SUBAPPLICATION Uebung_141_AX (* Übung zu DiagSetDTC: Drahtbruch 4-20 mA als DTC über DM1 *)
  (* Standard: 61499-2; Description: Copyright (c) 2026 Meisterschulen am Ostbahnhof This program and the accompanying materials are made available under the terms of the Eclipse Public License 2.0 which is available at https://www.eclipse.org/legal/epl-2.0/ SPDX-License-Identifier: EPL-2.0 *)
  (* Version 1.0, 2026-11-17, Franz Höpfinger, Meisterschulen am Ostbahnhof, initial API and implementation and/or initial documentation *)
  PACKAGE Uebungen;
  IMPORT Uebungen::const::Uebung_120_129::Filter::ADD_ALL_PASS;
  IMPORT Uebungen::const::Uebung_120_129::Filter::FLT_ALL_PASS;
  IMPORT Uebungen::const::Uebung_140_149::Diag::MV_DRAHTBRUCH;
  IMPORT Uebungen::const::Uebung_140_149::Diag::MV_OK;
  IMPORT Uebungen::const::Uebung_140_149::Diag::SPN_DRAHTBRUCH_AI6;
  IMPORT isobus::pgn::ISOUSERHOME_e::thisMember;
  IMPORT isobus::pgn::ISO_CAN_NODE::NODE1;
  IMPORT isobus::pgn::diag::FMI::CURRENT_LOW_OPEN_CIRCUIT;
  IMPORT logiBUS::io::AI::logiBUS_AI::AnalogInput_I6;
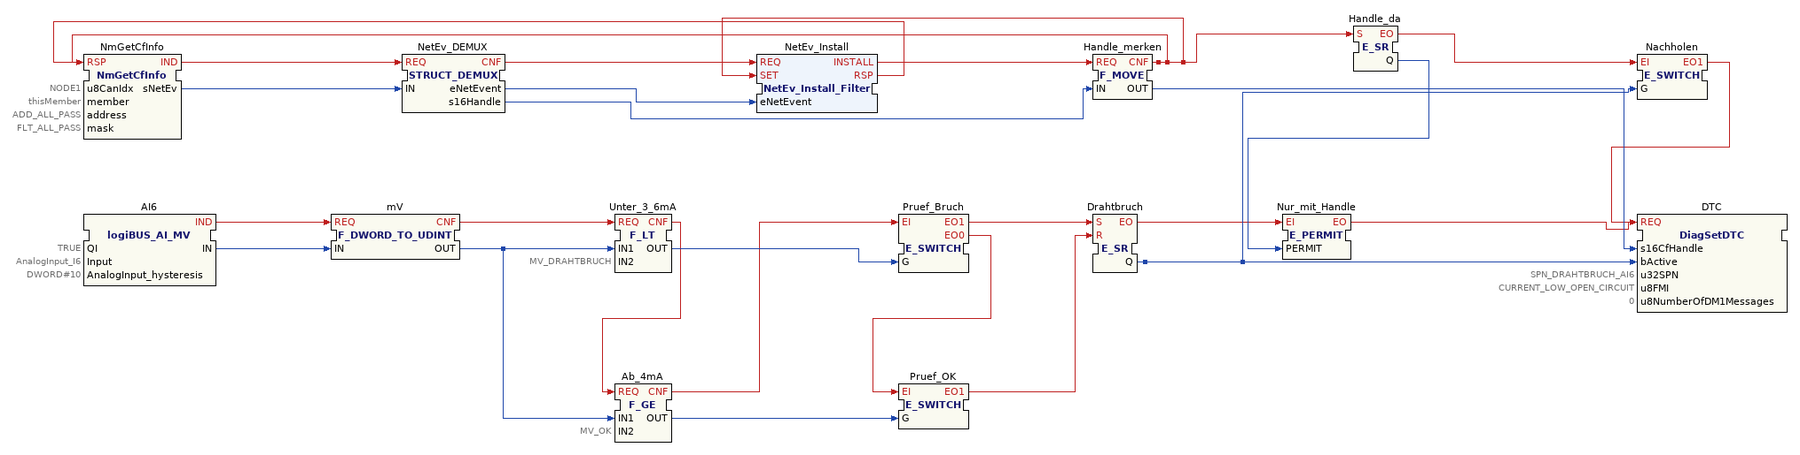
  (* Drahtbruch 4-20 mA an AI6 als DTC über DM1 (DiagSetDTC) Pin-mV unter 564 (3,6 mA) = Drahtbruch, wieder OK ab 626 (4 mA). Eigener CF-Handle aus NmGetCfInfo (thisMember, Active/NewAddress), RSP immer. DTC nur bei Zustandswechsel: SPN 520192, FMI 5, aktiv bis gelöscht. Test: Kabel ab = DM1 mit SPN 520192/FMI 5, jede Sekunde. Kabel dran = DTC inaktiv, in DM2, mit DM3 löschbar. Braucht Firmware ab LOGIBUS 96f591f2 (DM1) und isobus_pgn-ELF mit DiagSetDTC. *)
  FBS
    NmGetCfInfo : isobus::pgn::NmGetCfInfo(u8CanIdx := NODE1, member := thisMember, address := ADD_ALL_PASS, mask := FLT_ALL_PASS);
    NetEv_DEMUX : eclipse4diac::convert::STRUCT_DEMUX; {SET_ATTRIBUTE(StructuredType, isobus::pgn::ISONETEVENT_T)}
    Handle_merken : iec61131::selection::F_MOVE; (* eigener CF-Handle (s16Handle) *)
    Handle_da : iec61499::events::E_SR;
    Nachholen : iec61499::events::E_SWITCH; (* Drahtbruch schon vor dem Handle da: jetzt melden *)
    AI6 : logiBUS::io::AI::logiBUS_AI_MV(QI := TRUE, Input := AnalogInput_I6, AnalogInput_hysteresis := DWORD#10); (* mV am Pin, 4-20 mA über 491,2 Ohm *)
    mV : iec61131::conversion::F_DWORD_TO_UDINT;
    Unter_3_6mA : iec61131::comparison::F_LT(IN2 := MV_DRAHTBRUCH);
    Ab_4mA : iec61131::comparison::F_GE(IN2 := MV_OK);
    Pruef_Bruch : iec61499::events::E_SWITCH;
    Pruef_OK : iec61499::events::E_SWITCH;
    Drahtbruch : iec61499::events::E_SR; (* EO nur bei Zustandswechsel *)
    Nur_mit_Handle : iec61499::events::E_PERMIT;
    DTC : isobus::pgn::diag::DiagSetDTC(u32SPN := SPN_DRAHTBRUCH_AI6, u8FMI := CURRENT_LOW_OPEN_CIRCUIT, u8NumberOfDM1Messages := 0); (* DM1: SPN 520192, FMI 5 *)
  END_FBS
  SUBAPPS
    NetEv_Install : MyLib::sys::NetEv_Install_Filter;
  END_SUBAPPS
  EVENT_CONNECTIONS
    NmGetCfInfo.IND TO NetEv_DEMUX.REQ;
    NetEv_DEMUX.CNF TO NetEv_Install.REQ;
    NetEv_Install.INSTALL TO Handle_merken.REQ;
    NetEv_Install.RSP TO NmGetCfInfo.RSP;
    Handle_merken.CNF TO NetEv_Install.SET;
    Handle_merken.CNF TO Handle_da.S;
    Handle_merken.CNF TO NmGetCfInfo.RSP;
    Handle_da.EO TO Nachholen.EI;
    Nachholen.EO1 TO DTC.REQ;
    AI6.IND TO mV.REQ;
    mV.CNF TO Unter_3_6mA.REQ;
    Unter_3_6mA.CNF TO Ab_4mA.REQ;
    Ab_4mA.CNF TO Pruef_Bruch.EI;
    Pruef_Bruch.EO1 TO Drahtbruch.S;
    Pruef_Bruch.EO0 TO Pruef_OK.EI;
    Pruef_OK.EO1 TO Drahtbruch.R;
    Drahtbruch.EO TO Nur_mit_Handle.EI;
    Nur_mit_Handle.EO TO DTC.REQ;
  END_CONNECTIONS
  DATA_CONNECTIONS
    NmGetCfInfo.sNetEv TO NetEv_DEMUX.IN;
    NetEv_DEMUX.eNetEvent TO NetEv_Install.eNetEvent;
    NetEv_DEMUX.s16Handle TO Handle_merken.IN;
    Handle_merken.OUT TO DTC.s16CfHandle;
    Handle_da.Q TO Nur_mit_Handle.PERMIT;
    Drahtbruch.Q TO Nachholen.G;
    Drahtbruch.Q TO DTC.bActive;
    AI6.IN TO mV.IN;
    mV.OUT TO Unter_3_6mA.IN1;
    mV.OUT TO Ab_4mA.IN1;
    Unter_3_6mA.OUT TO Pruef_Bruch.G;
    Ab_4mA.OUT TO Pruef_OK.G;
  END_CONNECTIONS
END_SUBAPPLICATION
